(* PLC project Vn_fb_ctd, Beckhoff Automation GmbH TwinCAT PLC Control 3.5.13.21 *)
(* stored: creationDateTime 1970-01-01T00:00:00 *)

PROGRAM Vn_fb_ctd

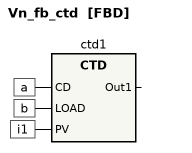
(* FBD diagram, written out as Structured Text *)
ctd1(CD := a, LOAD := b, PV := i1);
END_PROGRAM
